Staubli VAL3: cycle_Init.pgx

program cycle_Init()
begin
  //
  call Init()
  //
  call act:init()
  //
  call io:init()

  //  if !isPowered() and workingMode()==4
  //    enablePower()
  //    delay(1)
  //  endIf

end
